FUNCTION_BLOCK FB_LogRecordProcessor_Signoz EXTENDS FB_LogRecordProcessor_Simple
VAR_INPUT
END_VAR
VAR_OUTPUT
END_VAR
VAR
END_VAR

METHOD enrich
VAR_IN_OUT
	logRecord	: TcOtlp.FB_LogRecord;
END_VAR
IF logRecord.eventName <> 0 THEN
	logRecord.attributes.setStringAttribute('event.name', logRecord.eventName^.pString^);
END_IF
END_METHOD

END_FUNCTION_BLOCK

(* stored: Version 1.1.0.1
   POU FB_LogRecordProcessor_Signoz: Id {2571e0bd-c3f7-4d99-b45e-5120ce2bc3b4}, SpecialFunc None
   Method enrich: Id {91a52f0c-96a1-409b-81d1-5413c0486b5a} *)
